FUNCTION_BLOCK FB_LightTower_Control
VAR_INPUT
	ES_State		: BOOL;
	RunProcess1		: BOOL;
	RunProcess2		: BOOL;
	RunProcess3		: BOOL;
	ModeZone1		: E_ModeZone;
	ModeZone2		: E_ModeZone;
	ModeZone3		: E_ModeZone;
END_VAR

VAR_OUTPUT
	eLightTowerState		: E_LightTowerState;
END_VAR
VAR
END_VAR

IF ES_State THEN;
	IF stOper[ModeZone1].iActOperation=E_OperationButtons.ePauseAll 
	OR stOper[ModeZone2].iActOperation=E_OperationButtons.ePauseAll
	OR stOper[ModeZone3].iActOperation=E_OperationButtons.ePauseAll
	THEN;
		eLightTowerState:= E_LightTowerState.eYellow;
	ELSIF RunProcess1 OR RunProcess2 OR RunProcess3 THEN;
		eLightTowerState:= E_LightTowerState.eGreen;
	ELSE;
		eLightTowerState:= E_LightTowerState.eBlue;
	END_IF
	
ELSE;
	eLightTowerState:= E_LightTowerState.eRed;
END_IF

END_FUNCTION_BLOCK

(* stored: Version 1.1.0.1, ProductVersion 3.1.4024.15
   POU FB_LightTower_Control: Id {d4c40c7e-8f0e-41b4-947c-71820532771c}, SpecialFunc None *)
